// TIA Portal V20 export
// export: Created 2026-10-09T07:03:58.1914004Z, ExportSetting WithDefaults, DisplayName Totally Integrated Automation Portal, DisplayVersion V20, DisplayName TIA Portal Openness, DisplayVersion V20, DisplayName TIA Portal Teamcenter Gateway, DisplayVersion V20, DisplayName TIA Portal Version Control Interface, DisplayVersion V20, DisplayName SINAMICS Startdrive Advanced, DisplayVersion V20 SP1 Update 2, DisplayName SINAMICS Startdrive G110M, G120, G120C, G120D, G120P, G115D, DisplayVersion V20 SP1 Update 2, DisplayName SINAMICS Startdrive G130, G150, S120, S150, SINAMICS MV, G220, S200, S210, DisplayVersion V20 SP1 Update 2, DisplayName STEP 7 Professional, DisplayVersion V20, DisplayName STEP 7 Safety, DisplayVersion V20, DisplayName WinCC Basic/Comfort/Advanced, DisplayVersion V20, DisplayName WinCC Professional, DisplayVersion V20, DisplayName WinCC Unified, DisplayVersion V20
FUNCTION_BLOCK "FB_GRAPH_PressDemoAuto"   // FB100, GRAPH
VERSION : 0.1
// stored: AcknowledgeErrorsRequired true, AutoNumber true, GraphVersion 6.0, InitialValuesAcquisition false, IsIECCheckEnabled false, LanguageInNetworks LAD, LockOperatingMode false, PermanentILProcessingInMANMode false, SetENOAutomatically false, SkipSteps false, UDAEnableTagReadback false, WithAlarmHandling true
   // inherited from GRAPH_BASE
   VAR
      OFF_SQ_BASE : Bool;
   END_VAR
   VAR_INPUT
      OFF_SQ { ExternalAccessible := 'False'; ExternalVisible := 'False'; ExternalWritable := 'False'} : Bool := false;   // Turn sequence off
      INIT_SQ { ExternalAccessible := 'False'; ExternalVisible := 'False'; ExternalWritable := 'False'} : Bool := false;   // Set sequence to initial state
      ACK_EF { ExternalAccessible := 'False'; ExternalVisible := 'False'; ExternalWritable := 'False'} : Bool := false;   // Acknowledge all errors and faults
      S_PREV { ExternalAccessible := 'False'; ExternalVisible := 'False'; ExternalWritable := 'False'} : Bool := false;   // Output previous step in parameter S_NO
      S_NEXT { ExternalAccessible := 'False'; ExternalVisible := 'False'; ExternalWritable := 'False'} : Bool := false;   // Indicate next step in parameter S_NO
      SW_AUTO { ExternalAccessible := 'False'; ExternalVisible := 'False'; ExternalWritable := 'False'} : Bool := false;   // Automatic mode
      SW_TAP { ExternalAccessible := 'False'; ExternalVisible := 'False'; ExternalWritable := 'False'} : Bool := false;   // Semiautomatic/switch with transition
      SW_TOP { ExternalAccessible := 'False'; ExternalVisible := 'False'; ExternalWritable := 'False'} : Bool := false;   // Semiautomatic/ignore transition
      SW_MAN { ExternalAccessible := 'False'; ExternalVisible := 'False'; ExternalWritable := 'False'} : Bool := false;   // Manual mode
      S_SEL { ExternalAccessible := 'False'; ExternalVisible := 'False'; ExternalWritable := 'False'} : Int := 0;   // Select step to be output to S_NO
      S_ON { ExternalAccessible := 'False'; ExternalVisible := 'False'; ExternalWritable := 'False'} : Bool := false;   // Activate step indicated in S_NO
      S_OFF { ExternalAccessible := 'False'; ExternalVisible := 'False'; ExternalWritable := 'False'} : Bool := false;   // Disable step indicated in S_NO
      T_PUSH { ExternalAccessible := 'False'; ExternalVisible := 'False'; ExternalWritable := 'False'} : Bool := false;   // Enable transition to switch in semi automatic mode
      Run : BOOL;
      Reset : BOOL;
      OwnerIndex : DINT;
      Delta : TIME;
      TransferSettleTime : TIME;
      PartQuality : BOOL;
      RequireTwoHandStart : BOOL;
      SourcePath : String[80];
      PartPresent : BOOL;
      AirPressureOk : BOOL;
      TwoHandHeld : BOOL;
      StartPulse : BOOL;
      PressSettleTime : TIME;
   END_VAR
   VAR_OUTPUT
      S_NO { ExternalAccessible := 'False'; ExternalVisible := 'False'; ExternalWritable := 'False'} : Int := 0;   // Step number
      S_MORE { ExternalAccessible := 'False'; ExternalVisible := 'False'; ExternalWritable := 'False'} : Bool := false;   // More steps are available and can be shown in S_NO
      S_ACTIVE { ExternalAccessible := 'False'; ExternalVisible := 'False'; ExternalWritable := 'False'} : Bool := false;   // Step indicated in S_NO is active
      ERR_FLT { ExternalAccessible := 'False'; ExternalVisible := 'False'; ExternalWritable := 'False'} : Bool := false;   // Interlock or supervision group error
      AUTO_ON { ExternalAccessible := 'False'; ExternalVisible := 'False'; ExternalWritable := 'False'} : Bool := false;   // Automatic mode is active
      TAP_ON { ExternalAccessible := 'False'; ExternalVisible := 'False'; ExternalWritable := 'False'} : Bool := false;   // Semiautomatic mode/step with transition enabled
      TOP_ON { ExternalAccessible := 'False'; ExternalVisible := 'False'; ExternalWritable := 'False'} : Bool := false;   // Semiautomatic mode/ignore transition enabled
      MAN_ON { ExternalAccessible := 'False'; ExternalVisible := 'False'; ExternalWritable := 'False'} : Bool := false;   // Manual mode is active
   END_VAR
   VAR_IN_OUT
      PressRam : "FB_CylinderCM";
      Door : "FB_CylinderCM";
      PartSlide : "FB_CylinderCM";
      HostCore : "FRK_Core";
      HostUnit : "FRK_Unit";
      HostStatus : "ST_ModuleStatus";
      HostPart : "ST_PartContext";
      HostAlarmLog : "FRK_AlarmLog";
      Seq : "FRK_SequenceCtx";
      Row1 : "FRK_SequenceRow";
      Row2 : "FRK_SequenceRow";
      Row3 : "FRK_SequenceRow";
      Row4 : "FRK_SequenceRow";
      Row5 : "FRK_SequenceRow";
      Row6 : "FRK_SequenceRow";
      Row7 : "FRK_SequenceRow";
      Row8 : "FRK_SequenceRow";
      Row9 : "FRK_SequenceRow";
      Row10 : "FRK_SequenceRow";
      Row11 : "FRK_SequenceRow";
      Row12 : "FRK_SequenceRow";
      Row13 : "FRK_SequenceRow";
      Row14 : "FRK_SequenceRow";
      Row15 : "FRK_SequenceRow";
      Row16 : "FRK_SequenceRow";
      Ready1 { ExternalAccessible := 'False'; ExternalVisible := 'False'; ExternalWritable := 'False'} : BOOL;
      Ready2 { ExternalAccessible := 'False'; ExternalVisible := 'False'; ExternalWritable := 'False'} : BOOL;
      Ready3 { ExternalAccessible := 'False'; ExternalVisible := 'False'; ExternalWritable := 'False'} : BOOL;
      Ready4 { ExternalAccessible := 'False'; ExternalVisible := 'False'; ExternalWritable := 'False'} : BOOL;
      Ready5 { ExternalAccessible := 'False'; ExternalVisible := 'False'; ExternalWritable := 'False'} : BOOL;
      Cycle : "ST_PressDemoCycle";
      LoadDone { ExternalAccessible := 'False'; ExternalVisible := 'False'; ExternalWritable := 'False'} : BOOL;
      Branch1 : "FRK_SequenceCtx";
      Branch2 : "FRK_SequenceCtx";
      Row17 : "FRK_SequenceRow";
      Row18 : "FRK_SequenceRow";
      Row19 : "FRK_SequenceRow";
   END_VAR
BEGIN
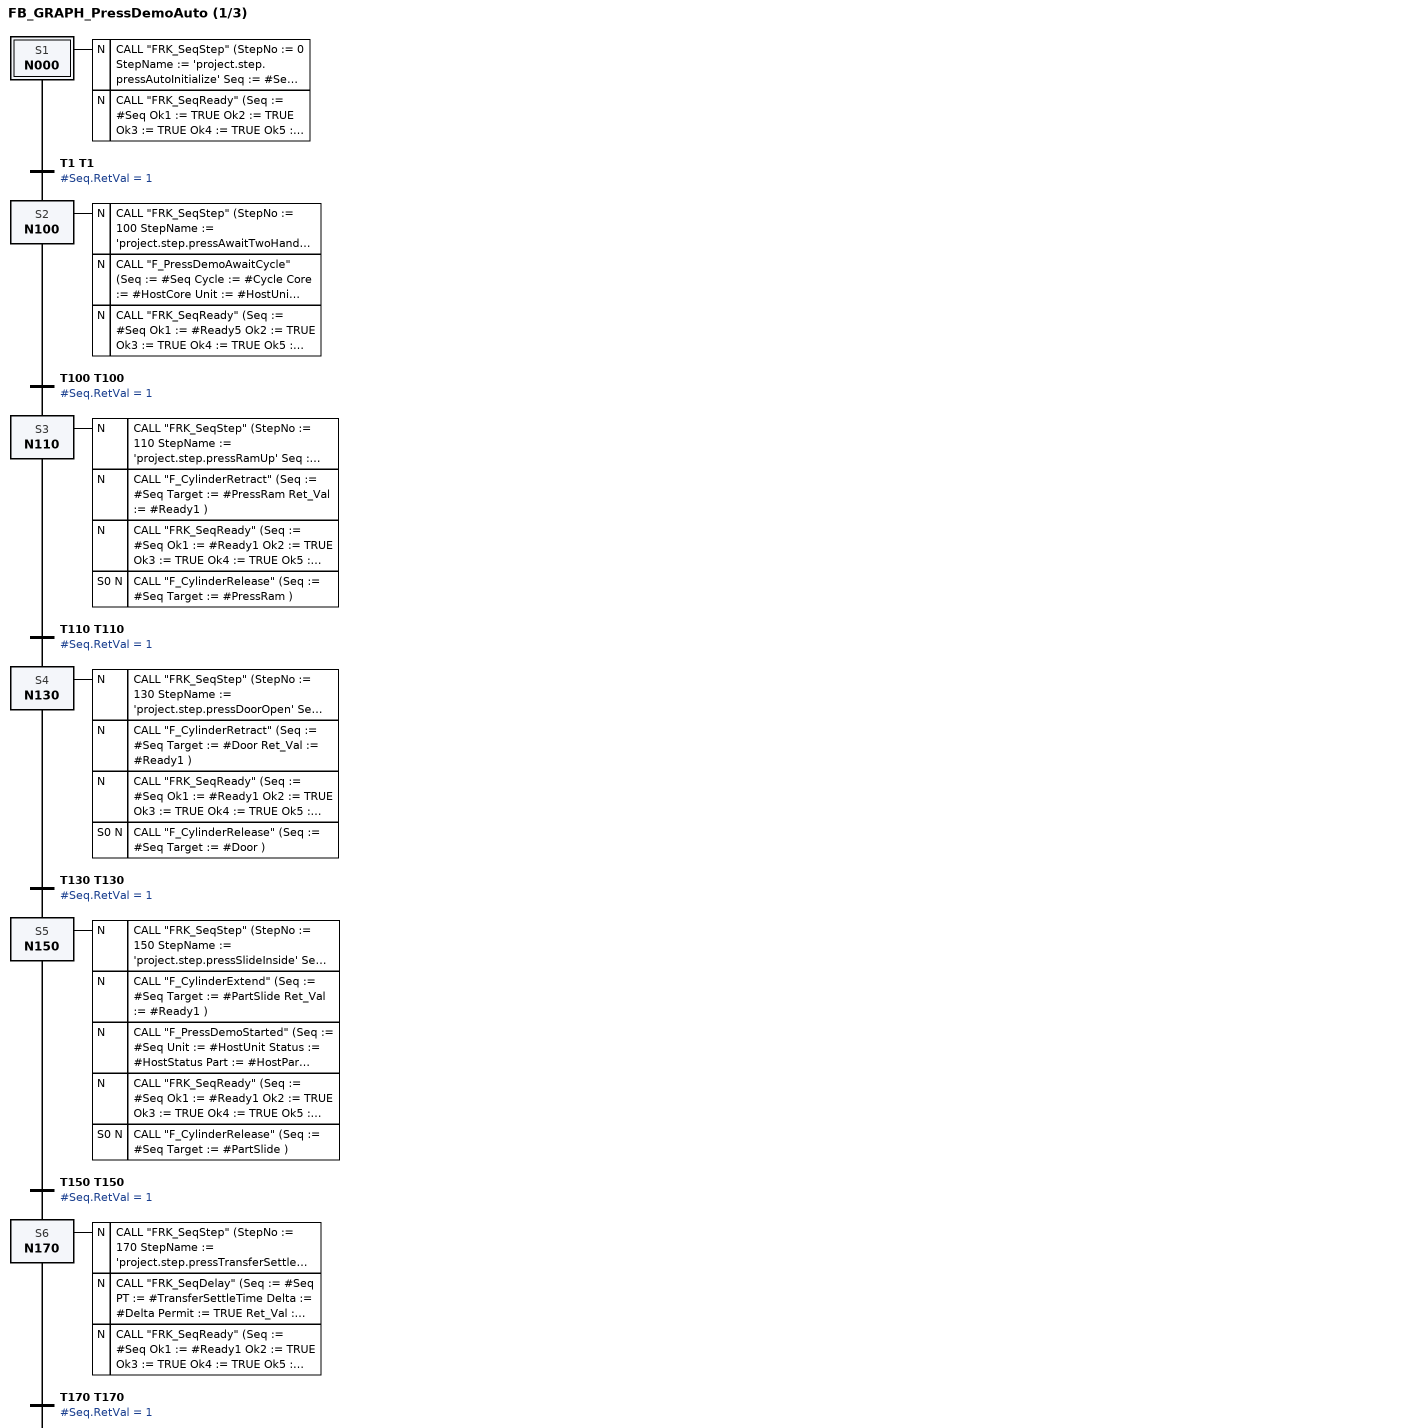
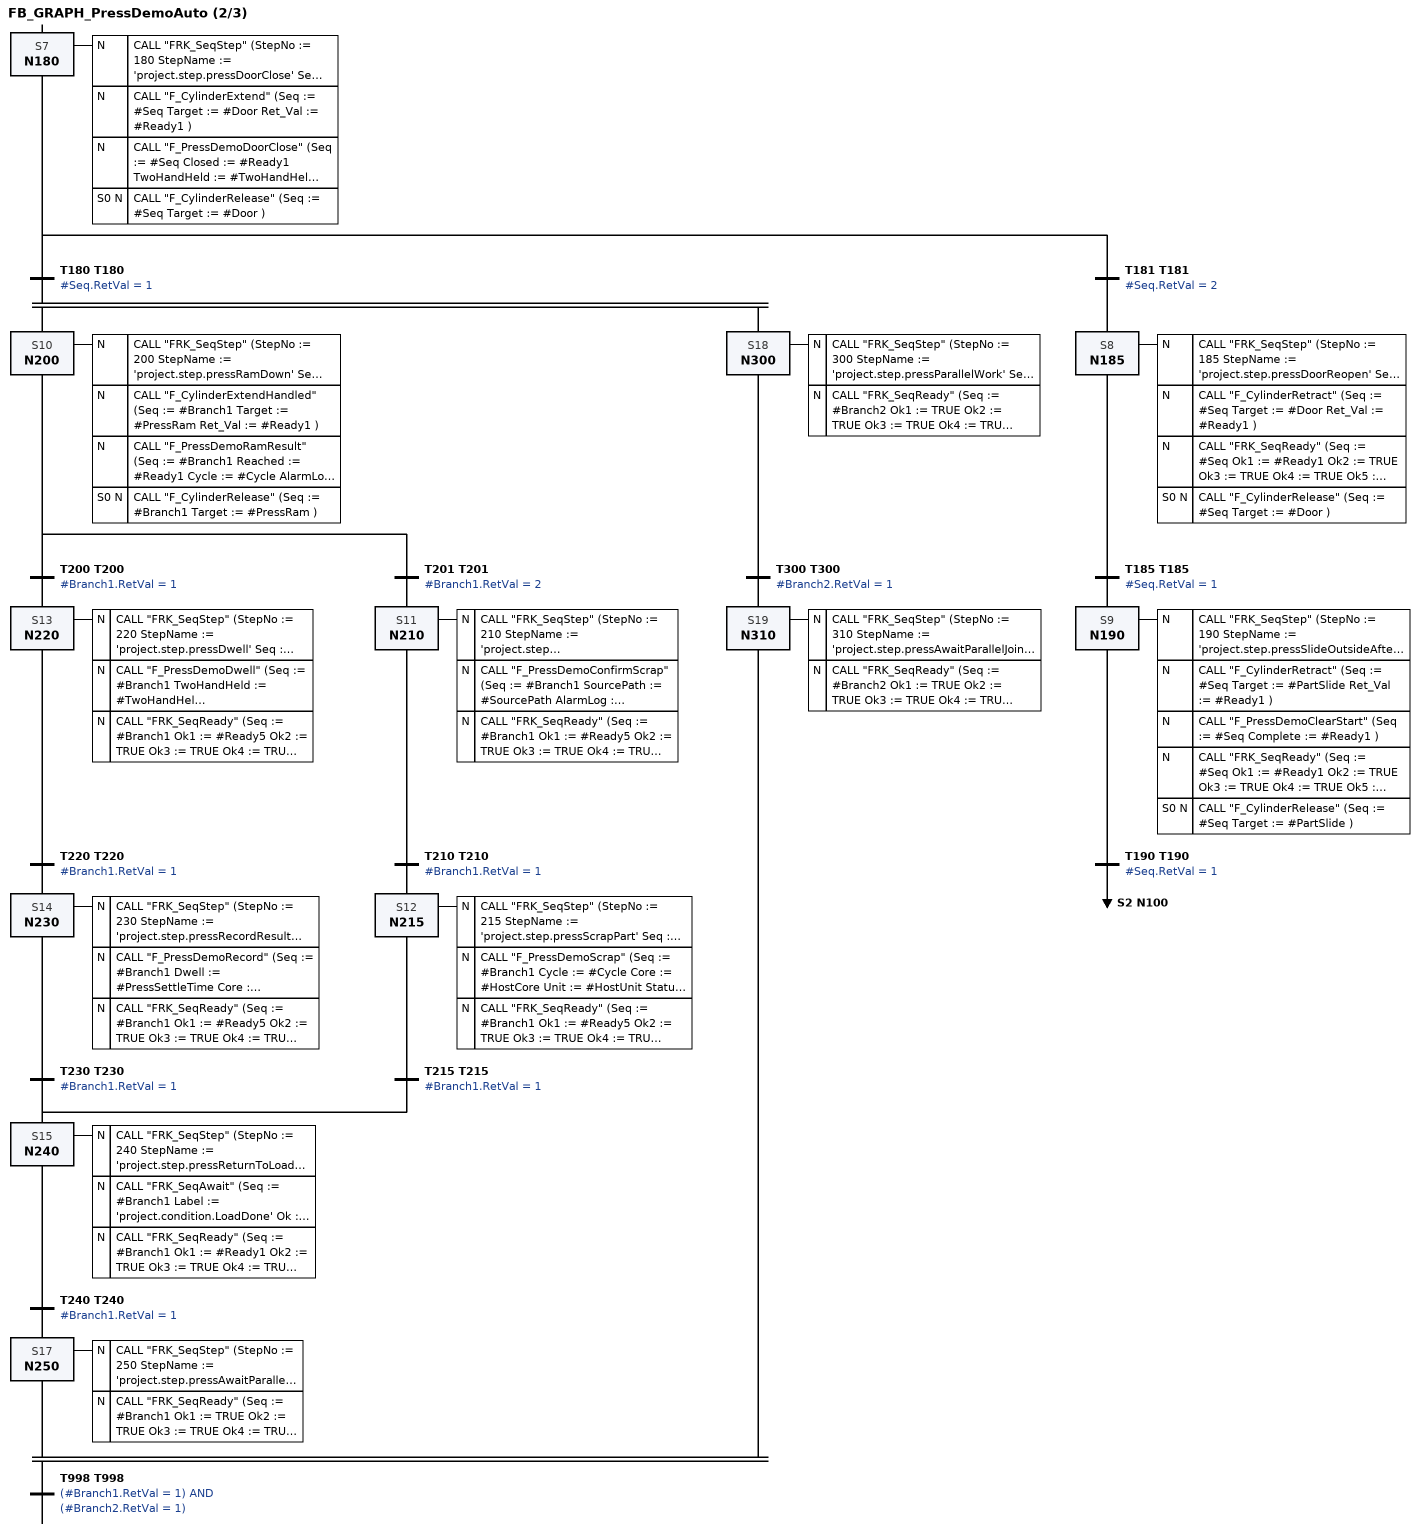
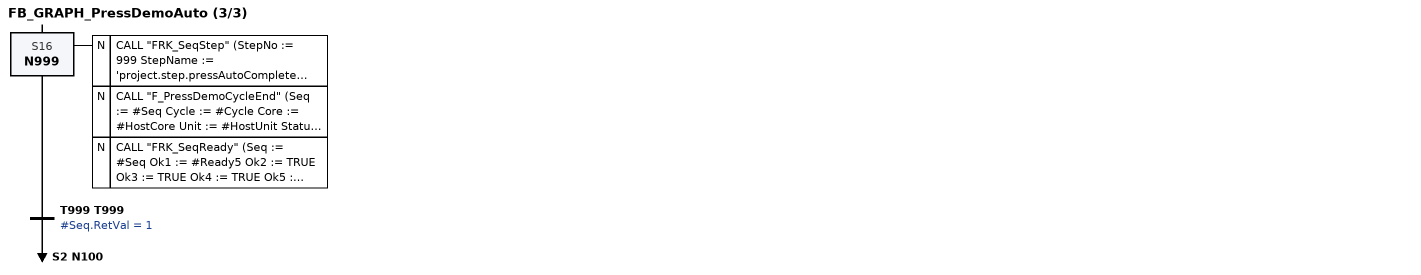
   // sequencer 1
   INITIAL_STEP N000:   // S1, max time T#10S, warning time T#7S
              N    CALL "FRK_SeqStep" 
                   (StepNo := 0
                   StepName := 'project.step.pressAutoInitialize'
                   Seq := #Seq
                   Row := #Row1
                   )
              N    CALL "FRK_SeqReady" 
                   (Seq := #Seq
                   Ok1 := TRUE
                   Ok2 := TRUE
                   Ok3 := TRUE
                   Ok4 := TRUE
                   Ok5 := TRUE
                   )
   END_STEP
   TRANSITION T1 FROM N000 TO N100   // T1
      := #Seq.RetVal = 1;
   END_TRANSITION
   STEP N100:   // S2, max time T#10S, warning time T#7S
              N    CALL "FRK_SeqStep" 
                   (StepNo := 100
                   StepName := 'project.step.pressAwaitTwoHand'
                   Seq := #Seq
                   Row := #Row2
                   )
              N    CALL "F_PressDemoAwaitCycle" 
                   (Seq := #Seq
                   Cycle := #Cycle
                   Core := #HostCore
                   Unit := #HostUnit
                   Status := #HostStatus
                   Part := #HostPart
                   AlarmLog := #HostAlarmLog
                   PartPresent := #PartPresent
                   PartQuality := #PartQuality
                   AirPressureOk := #AirPressureOk
                   RequireTwoHandStart := #RequireTwoHandStart
                   Ret_Val := #Ready5
                   )
              N    CALL "FRK_SeqReady" 
                   (Seq := #Seq
                   Ok1 := #Ready5
                   Ok2 := TRUE
                   Ok3 := TRUE
                   Ok4 := TRUE
                   Ok5 := TRUE
                   )
   END_STEP
   TRANSITION T100 FROM N100 TO N110   // T100
      := #Seq.RetVal = 1;
   END_TRANSITION
   STEP N110:   // S3, max time T#10S, warning time T#7S
              N    CALL "FRK_SeqStep" 
                   (StepNo := 110
                   StepName := 'project.step.pressRamUp'
                   Seq := #Seq
                   Row := #Row3
                   )
              N    CALL "F_CylinderRetract" 
                   (Seq := #Seq
                   Target := #PressRam
                   Ret_Val := #Ready1
                   )
              N    CALL "FRK_SeqReady" 
                   (Seq := #Seq
                   Ok1 := #Ready1
                   Ok2 := TRUE
                   Ok3 := TRUE
                   Ok4 := TRUE
                   Ok5 := TRUE
                   )
          S0  N    CALL "F_CylinderRelease" 
                   (Seq := #Seq
                   Target := #PressRam
                   )
   END_STEP
   TRANSITION T110 FROM N110 TO N130   // T110
      := #Seq.RetVal = 1;
   END_TRANSITION
   STEP N130:   // S4, max time T#10S, warning time T#7S
              N    CALL "FRK_SeqStep" 
                   (StepNo := 130
                   StepName := 'project.step.pressDoorOpen'
                   Seq := #Seq
                   Row := #Row4
                   )
              N    CALL "F_CylinderRetract" 
                   (Seq := #Seq
                   Target := #Door
                   Ret_Val := #Ready1
                   )
              N    CALL "FRK_SeqReady" 
                   (Seq := #Seq
                   Ok1 := #Ready1
                   Ok2 := TRUE
                   Ok3 := TRUE
                   Ok4 := TRUE
                   Ok5 := TRUE
                   )
          S0  N    CALL "F_CylinderRelease" 
                   (Seq := #Seq
                   Target := #Door
                   )
   END_STEP
   TRANSITION T130 FROM N130 TO N150   // T130
      := #Seq.RetVal = 1;
   END_TRANSITION
   STEP N150:   // S5, max time T#10S, warning time T#7S
              N    CALL "FRK_SeqStep" 
                   (StepNo := 150
                   StepName := 'project.step.pressSlideInside'
                   Seq := #Seq
                   Row := #Row5
                   )
              N    CALL "F_CylinderExtend" 
                   (Seq := #Seq
                   Target := #PartSlide
                   Ret_Val := #Ready1
                   )
              N    CALL "F_PressDemoStarted" 
                   (Seq := #Seq
                   Unit := #HostUnit
                   Status := #HostStatus
                   Part := #HostPart
                   AlarmLog := #HostAlarmLog
                   )
              N    CALL "FRK_SeqReady" 
                   (Seq := #Seq
                   Ok1 := #Ready1
                   Ok2 := TRUE
                   Ok3 := TRUE
                   Ok4 := TRUE
                   Ok5 := TRUE
                   )
          S0  N    CALL "F_CylinderRelease" 
                   (Seq := #Seq
                   Target := #PartSlide
                   )
   END_STEP
   TRANSITION T150 FROM N150 TO N170   // T150
      := #Seq.RetVal = 1;
   END_TRANSITION
   STEP N170:   // S6, max time T#10S, warning time T#7S
              N    CALL "FRK_SeqStep" 
                   (StepNo := 170
                   StepName := 'project.step.pressTransferSettle'
                   Seq := #Seq
                   Row := #Row6
                   )
              N    CALL "FRK_SeqDelay" 
                   (Seq := #Seq
                   PT := #TransferSettleTime
                   Delta := #Delta
                   Permit := TRUE
                   Ret_Val := #Ready1
                   )
              N    CALL "FRK_SeqReady" 
                   (Seq := #Seq
                   Ok1 := #Ready1
                   Ok2 := TRUE
                   Ok3 := TRUE
                   Ok4 := TRUE
                   Ok5 := TRUE
                   )
   END_STEP
   TRANSITION T170 FROM N170 TO N180   // T170
      := #Seq.RetVal = 1;
   END_TRANSITION
   STEP N180:   // S7, max time T#10S, warning time T#7S
              N    CALL "FRK_SeqStep" 
                   (StepNo := 180
                   StepName := 'project.step.pressDoorClose'
                   Seq := #Seq
                   Row := #Row7
                   )
              N    CALL "F_CylinderExtend" 
                   (Seq := #Seq
                   Target := #Door
                   Ret_Val := #Ready1
                   )
              N    CALL "F_PressDemoDoorClose" 
                   (Seq := #Seq
                   Closed := #Ready1
                   TwoHandHeld := #TwoHandHeld
                   RequireTwoHandStart := #RequireTwoHandStart
                   SourcePath := #SourcePath
                   AlarmLog := #HostAlarmLog
                   )
          S0  N    CALL "F_CylinderRelease" 
                   (Seq := #Seq
                   Target := #Door
                   )
   END_STEP
   TRANSITION T180 FROM N180 TO (N200, N300)   // T180
      := #Seq.RetVal = 1;
   END_TRANSITION
   TRANSITION T181 FROM N180 TO N185   // T181
      := #Seq.RetVal = 2;
   END_TRANSITION
   STEP N185:   // S8, max time T#10S, warning time T#7S
              N    CALL "FRK_SeqStep" 
                   (StepNo := 185
                   StepName := 'project.step.pressDoorReopen'
                   Seq := #Seq
                   Row := #Row8
                   )
              N    CALL "F_CylinderRetract" 
                   (Seq := #Seq
                   Target := #Door
                   Ret_Val := #Ready1
                   )
              N    CALL "FRK_SeqReady" 
                   (Seq := #Seq
                   Ok1 := #Ready1
                   Ok2 := TRUE
                   Ok3 := TRUE
                   Ok4 := TRUE
                   Ok5 := TRUE
                   )
          S0  N    CALL "F_CylinderRelease" 
                   (Seq := #Seq
                   Target := #Door
                   )
   END_STEP
   TRANSITION T185 FROM N185 TO N190   // T185
      := #Seq.RetVal = 1;
   END_TRANSITION
   STEP N190:   // S9, max time T#10S, warning time T#7S
              N    CALL "FRK_SeqStep" 
                   (StepNo := 190
                   StepName := 'project.step.pressSlideOutsideAfterAbort'
                   Seq := #Seq
                   Row := #Row9
                   )
              N    CALL "F_CylinderRetract" 
                   (Seq := #Seq
                   Target := #PartSlide
                   Ret_Val := #Ready1
                   )
              N    CALL "F_PressDemoClearStart" 
                   (Seq := #Seq
                   Complete := #Ready1
                   )
              N    CALL "FRK_SeqReady" 
                   (Seq := #Seq
                   Ok1 := #Ready1
                   Ok2 := TRUE
                   Ok3 := TRUE
                   Ok4 := TRUE
                   Ok5 := TRUE
                   )
          S0  N    CALL "F_CylinderRelease" 
                   (Seq := #Seq
                   Target := #PartSlide
                   )
   END_STEP
   TRANSITION T190 FROM N190 TO N100   // T190, jump
      := #Seq.RetVal = 1;
   END_TRANSITION
   STEP N200:   // S10, max time T#10S, warning time T#7S
              N    CALL "FRK_SeqStep" 
                   (StepNo := 200
                   StepName := 'project.step.pressRamDown'
                   Seq := #Branch1
                   Row := #Row10
                   )
              N    CALL "F_CylinderExtendHandled" 
                   (Seq := #Branch1
                   Target := #PressRam
                   Ret_Val := #Ready1
                   )
              N    CALL "F_PressDemoRamResult" 
                   (Seq := #Branch1
                   Reached := #Ready1
                   Cycle := #Cycle
                   AlarmLog := #HostAlarmLog
                   )
          S0  N    CALL "F_CylinderRelease" 
                   (Seq := #Branch1
                   Target := #PressRam
                   )
   END_STEP
   TRANSITION T200 FROM N200 TO N220   // T200
      := #Branch1.RetVal = 1;
   END_TRANSITION
   TRANSITION T201 FROM N200 TO N210   // T201
      := #Branch1.RetVal = 2;
   END_TRANSITION
   STEP N210:   // S11, max time T#10S, warning time T#7S
              N    CALL "FRK_SeqStep" 
                   (StepNo := 210
                   StepName := 'project.step.pressNotReachedConfirm'
                   Seq := #Branch1
                   Row := #Row11
                   )
              N    CALL "F_PressDemoConfirmScrap" 
                   (Seq := #Branch1
                   SourcePath := #SourcePath
                   AlarmLog := #HostAlarmLog
                   Ret_Val := #Ready5
                   )
              N    CALL "FRK_SeqReady" 
                   (Seq := #Branch1
                   Ok1 := #Ready5
                   Ok2 := TRUE
                   Ok3 := TRUE
                   Ok4 := TRUE
                   Ok5 := TRUE
                   )
   END_STEP
   TRANSITION T210 FROM N210 TO N215   // T210
      := #Branch1.RetVal = 1;
   END_TRANSITION
   STEP N215:   // S12, max time T#10S, warning time T#7S
              N    CALL "FRK_SeqStep" 
                   (StepNo := 215
                   StepName := 'project.step.pressScrapPart'
                   Seq := #Branch1
                   Row := #Row12
                   )
              N    CALL "F_PressDemoScrap" 
                   (Seq := #Branch1
                   Cycle := #Cycle
                   Core := #HostCore
                   Unit := #HostUnit
                   Status := #HostStatus
                   Part := #HostPart
                   AlarmLog := #HostAlarmLog
                   Ret_Val := #Ready5
                   )
              N    CALL "FRK_SeqReady" 
                   (Seq := #Branch1
                   Ok1 := #Ready5
                   Ok2 := TRUE
                   Ok3 := TRUE
                   Ok4 := TRUE
                   Ok5 := TRUE
                   )
   END_STEP
   TRANSITION T215 FROM N215 TO N240   // T215
      := #Branch1.RetVal = 1;
   END_TRANSITION
   STEP N220:   // S13, max time T#10S, warning time T#7S
              N    CALL "FRK_SeqStep" 
                   (StepNo := 220
                   StepName := 'project.step.pressDwell'
                   Seq := #Branch1
                   Row := #Row13
                   )
              N    CALL "F_PressDemoDwell" 
                   (Seq := #Branch1
                   TwoHandHeld := #TwoHandHeld
                   RequireTwoHandStart := #RequireTwoHandStart
                   PT := #PressSettleTime
                   Delta := #Delta
                   PressRam := #PressRam
                   Ret_Val := #Ready5
                   )
              N    CALL "FRK_SeqReady" 
                   (Seq := #Branch1
                   Ok1 := #Ready5
                   Ok2 := TRUE
                   Ok3 := TRUE
                   Ok4 := TRUE
                   Ok5 := TRUE
                   )
   END_STEP
   TRANSITION T220 FROM N220 TO N230   // T220
      := #Branch1.RetVal = 1;
   END_TRANSITION
   STEP N230:   // S14, max time T#10S, warning time T#7S
              N    CALL "FRK_SeqStep" 
                   (StepNo := 230
                   StepName := 'project.step.pressRecordResult'
                   Seq := #Branch1
                   Row := #Row14
                   )
              N    CALL "F_PressDemoRecord" 
                   (Seq := #Branch1
                   Dwell := #PressSettleTime
                   Core := #HostCore
                   Status := #HostStatus
                   Part := #HostPart
                   Ret_Val := #Ready5
                   )
              N    CALL "FRK_SeqReady" 
                   (Seq := #Branch1
                   Ok1 := #Ready5
                   Ok2 := TRUE
                   Ok3 := TRUE
                   Ok4 := TRUE
                   Ok5 := TRUE
                   )
   END_STEP
   TRANSITION T230 FROM N230 TO N240   // T230
      := #Branch1.RetVal = 1;
   END_TRANSITION
   STEP N240:   // S15, max time T#10S, warning time T#7S
              N    CALL "FRK_SeqStep" 
                   (StepNo := 240
                   StepName := 'project.step.pressReturnToLoad'
                   Seq := #Branch1
                   Row := #Row15
                   )
              N    CALL "FRK_SeqAwait" 
                   (Seq := #Branch1
                   Label := 'project.condition.LoadDone'
                   Ok := #LoadDone
                   Ret_Val := #Ready1
                   )
              N    CALL "FRK_SeqReady" 
                   (Seq := #Branch1
                   Ok1 := #Ready1
                   Ok2 := TRUE
                   Ok3 := TRUE
                   Ok4 := TRUE
                   Ok5 := TRUE
                   )
   END_STEP
   TRANSITION T240 FROM N240 TO N250   // T240
      := #Branch1.RetVal = 1;
   END_TRANSITION
   STEP N999:   // S16, max time T#10S, warning time T#7S
              N    CALL "FRK_SeqStep" 
                   (StepNo := 999
                   StepName := 'project.step.pressAutoComplete'
                   Seq := #Seq
                   Row := #Row16
                   )
              N    CALL "F_PressDemoCycleEnd" 
                   (Seq := #Seq
                   Cycle := #Cycle
                   Core := #HostCore
                   Unit := #HostUnit
                   Status := #HostStatus
                   Part := #HostPart
                   AlarmLog := #HostAlarmLog
                   Ret_Val := #Ready5
                   )
              N    CALL "FRK_SeqReady" 
                   (Seq := #Seq
                   Ok1 := #Ready5
                   Ok2 := TRUE
                   Ok3 := TRUE
                   Ok4 := TRUE
                   Ok5 := TRUE
                   )
   END_STEP
   TRANSITION T999 FROM N999 TO N100   // T999, jump
      := #Seq.RetVal = 1;
   END_TRANSITION
   STEP N250:   // S17, max time T#10S, warning time T#7S
              N    CALL "FRK_SeqStep" 
                   (StepNo := 250
                   StepName := 'project.step.pressAwaitParallelBranch'
                   Seq := #Branch1
                   Row := #Row17
                   )
              N    CALL "FRK_SeqReady" 
                   (Seq := #Branch1
                   Ok1 := TRUE
                   Ok2 := TRUE
                   Ok3 := TRUE
                   Ok4 := TRUE
                   Ok5 := TRUE
                   )
   END_STEP
   STEP N300:   // S18, max time T#10S, warning time T#7S
              N    CALL "FRK_SeqStep" 
                   (StepNo := 300
                   StepName := 'project.step.pressParallelWork'
                   Seq := #Branch2
                   Row := #Row18
                   )
              N    CALL "FRK_SeqReady" 
                   (Seq := #Branch2
                   Ok1 := TRUE
                   Ok2 := TRUE
                   Ok3 := TRUE
                   Ok4 := TRUE
                   Ok5 := TRUE
                   )
   END_STEP
   TRANSITION T300 FROM N300 TO N310   // T300
      := #Branch2.RetVal = 1;
   END_TRANSITION
   STEP N310:   // S19, max time T#10S, warning time T#7S
              N    CALL "FRK_SeqStep" 
                   (StepNo := 310
                   StepName := 'project.step.pressAwaitParallelJoin'
                   Seq := #Branch2
                   Row := #Row19
                   )
              N    CALL "FRK_SeqReady" 
                   (Seq := #Branch2
                   Ok1 := TRUE
                   Ok2 := TRUE
                   Ok3 := TRUE
                   Ok4 := TRUE
                   Ok5 := TRUE
                   )
   END_STEP
   TRANSITION T998 FROM (N250, N310) TO N999   // T998
      := (#Branch1.RetVal = 1) AND (#Branch2.RetVal = 1);
   END_TRANSITION
END_FUNCTION_BLOCK
